TYPE eLightCmdSource :
(
    NONE,
    SWITCH,
    HA,
    SCHEDULER,
	ROOM
);
END_TYPE

(* stored: Version 1.1.0.1
   DUT eLightCmdSource: Id {eabe1d87-a0b8-4beb-aa3e-3cd1c99bbe9f} *)
